FUNCTION_BLOCK Grade_Inovaisa (* Grade mecanizada do painel Vibropac com os niveis montante, jusante e diferencial - HidrycoLib *)
  (* Standard: 61499-2 *)
  (* Version 1.1, 11/11/2026, Hidryco, Hidryco, 1.1: sensores com cfgSkid = TRUE (niveis ja escalados no painel; sem ajuste de escala na IHM). 1.0: uma grade do gradeamento (padrao Grade_Equipamentos do legado): SensorMontante, SensorJusante, SensorDiferencial (Sensor_Generico por comunicacao, %) e Grade_Mecanizada_Inovaisa1 (Motor_Inovaisa com reverso e sobretorque). Os niveis chegam do processo e vao aos sensores por symlink ${PATH}SensorX.stsEntrada / stsFalhaComunicacao. *)
  PACKAGE Hidryco.HidrycoLib;
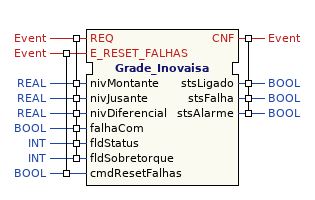
  EVENT_INPUT
    REQ WITH nivMontante, nivJusante, nivDiferencial, falhaCom, fldStatus, fldSobretorque; (* Leitura do painel (pelo processo) *)
    E_RESET_FALHAS WITH cmdResetFalhas; (* Reset dos sensores e reconhecimento dos alarmes (com cmdResetFalhas = TRUE) *)
  END_EVENT
  EVENT_OUTPUT
    CNF WITH stsLigado, stsFalha, stsAlarme; (* Status da grade (na mudanca) *)
  END_EVENT
  VAR_INPUT
    nivMontante : REAL; (* Nivel montante (%) *)
    nivJusante : REAL; (* Nivel jusante (%) *)
    nivDiferencial : REAL; (* Nivel diferencial (%) *)
    falhaCom : BOOL; (* Sem comunicacao com o painel *)
    fldStatus : INT; (* Registro de status da grade (4007/4008) *)
    fldSobretorque : INT; (* Registro do sobretorque (4010/4011) *)
    cmdResetFalhas : BOOL; (* TRUE = reset (com o evento E_RESET_FALHAS) *)
  END_VAR
  VAR_OUTPUT
    stsLigado : BOOL; (* Grade funcionando *)
    stsFalha : BOOL; (* Grade em falha *)
    stsAlarme : BOOL; (* Falha ou sobretorque *)
  END_VAR
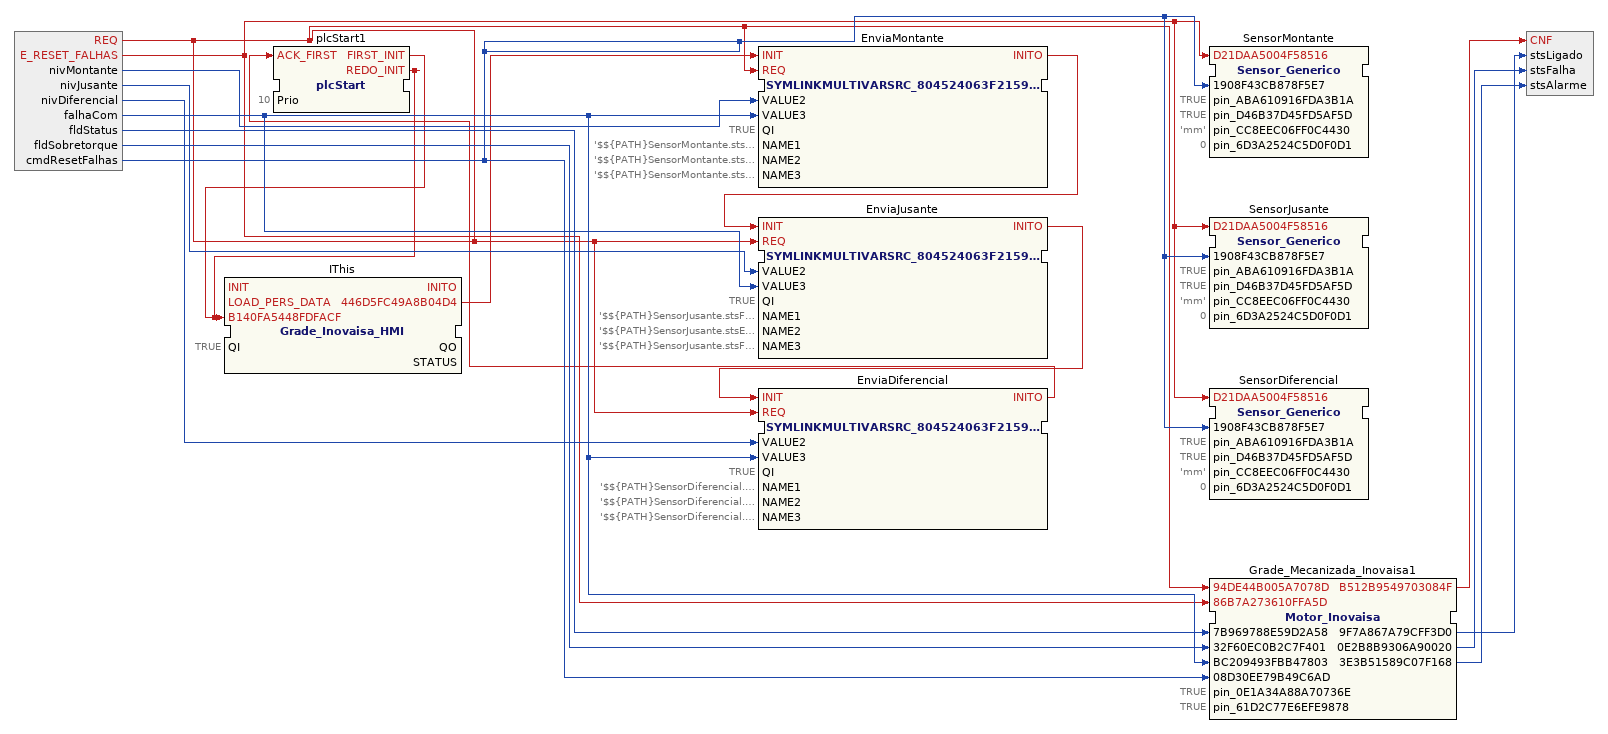
  FBS
    IThis : Grade_Inovaisa_HMI(QI := TRUE);
    plcStart1 : plcStart(Prio := 10);
    SensorMontante : Sensor_Generico(pin_ABA610916FDA3B1A := TRUE, pin_D46B37D45FD5AF5D := TRUE, pin_CC8EEC06FF0C4430 := 'mm', pin_6D3A2524C5D0F0D1 := 0);
    EnviaMontante : SYMLINKMULTIVARSRC_804524063F215924(QI := TRUE, NAME1 := '$${PATH}SensorMontante.stsFalhaSensor', NAME2 := '$${PATH}SensorMontante.stsEntrada', NAME3 := '$${PATH}SensorMontante.stsFalhaComunicacao'); {SET_ATTRIBUTE(Configuration.GenericFBType.InterfaceParams, Runtime.System#I:=3;VALUE${I$}:BOOL,REAL,BOOL)}
    SensorJusante : Sensor_Generico(pin_ABA610916FDA3B1A := TRUE, pin_D46B37D45FD5AF5D := TRUE, pin_CC8EEC06FF0C4430 := 'mm', pin_6D3A2524C5D0F0D1 := 0);
    EnviaJusante : SYMLINKMULTIVARSRC_804524063F215924(QI := TRUE, NAME1 := '$${PATH}SensorJusante.stsFalhaSensor', NAME2 := '$${PATH}SensorJusante.stsEntrada', NAME3 := '$${PATH}SensorJusante.stsFalhaComunicacao'); {SET_ATTRIBUTE(Configuration.GenericFBType.InterfaceParams, Runtime.System#I:=3;VALUE${I$}:BOOL,REAL,BOOL)}
    SensorDiferencial : Sensor_Generico(pin_ABA610916FDA3B1A := TRUE, pin_D46B37D45FD5AF5D := TRUE, pin_CC8EEC06FF0C4430 := 'mm', pin_6D3A2524C5D0F0D1 := 0);
    EnviaDiferencial : SYMLINKMULTIVARSRC_804524063F215924(QI := TRUE, NAME1 := '$${PATH}SensorDiferencial.stsFalhaSensor', NAME2 := '$${PATH}SensorDiferencial.stsEntrada', NAME3 := '$${PATH}SensorDiferencial.stsFalhaComunicacao'); {SET_ATTRIBUTE(Configuration.GenericFBType.InterfaceParams, Runtime.System#I:=3;VALUE${I$}:BOOL,REAL,BOOL)}
    Grade_Mecanizada_Inovaisa1 : Motor_Inovaisa(pin_0E1A34A88A70736E := TRUE, pin_61D2C77E6EFE9878 := TRUE);
  END_FBS
  EVENT_CONNECTIONS
    plcStart1.FIRST_INIT TO IThis.B140FA5448FDFACF;
    plcStart1.REDO_INIT TO IThis.B140FA5448FDFACF;
    IThis.446D5FC49A8B04D4 TO EnviaMontante.INIT;
    EnviaMontante.INITO TO EnviaJusante.INIT;
    EnviaJusante.INITO TO EnviaDiferencial.INIT;
    EnviaDiferencial.INITO TO plcStart1.ACK_FIRST;
    REQ TO EnviaMontante.REQ;
    E_RESET_FALHAS TO SensorMontante.D21DAA5004F58516;
    REQ TO EnviaJusante.REQ;
    E_RESET_FALHAS TO SensorJusante.D21DAA5004F58516;
    REQ TO EnviaDiferencial.REQ;
    E_RESET_FALHAS TO SensorDiferencial.D21DAA5004F58516;
    REQ TO Grade_Mecanizada_Inovaisa1.94DE44B005A7078D;
    E_RESET_FALHAS TO Grade_Mecanizada_Inovaisa1.86B7A273610FFA5D;
    Grade_Mecanizada_Inovaisa1.B512B9549703084F TO CNF;
  END_CONNECTIONS
  DATA_CONNECTIONS
    nivMontante TO EnviaMontante.VALUE2;
    falhaCom TO EnviaMontante.VALUE3;
    cmdResetFalhas TO SensorMontante.1908F43CB878F5E7;
    nivJusante TO EnviaJusante.VALUE2;
    falhaCom TO EnviaJusante.VALUE3;
    cmdResetFalhas TO SensorJusante.1908F43CB878F5E7;
    nivDiferencial TO EnviaDiferencial.VALUE2;
    falhaCom TO EnviaDiferencial.VALUE3;
    cmdResetFalhas TO SensorDiferencial.1908F43CB878F5E7;
    fldStatus TO Grade_Mecanizada_Inovaisa1.7B969788E59D2A58;
    fldSobretorque TO Grade_Mecanizada_Inovaisa1.32F60EC0B2C7F401;
    falhaCom TO Grade_Mecanizada_Inovaisa1.BC209493FBB47803;
    cmdResetFalhas TO Grade_Mecanizada_Inovaisa1.08D30EE79B49C6AD;
    Grade_Mecanizada_Inovaisa1.9F7A867A79CFF3D0 TO stsLigado;
    Grade_Mecanizada_Inovaisa1.0E2B8B9306A90020 TO stsFalha;
    Grade_Mecanizada_Inovaisa1.3E3B51589C07F168 TO stsAlarme;
  END_CONNECTIONS
END_FUNCTION_BLOCK
